// TIA Portal V15.1 export
// export: Created 2000-01-01T00:00:00.0000000Z, ExportSetting None
FUNCTION "FC_Rung" : Void   // FC42, LAD
{ S7_Optimized_Access := 'TRUE' }
   VAR_INPUT
      Local : Int;
   END_VAR
BEGIN

REGION Network 1
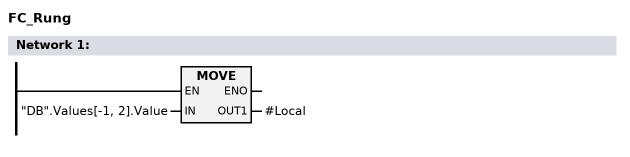
   RUNG wire#powerrail
      Move(in := "DB".Values[-1, 2].Value, out1 => #Local)
   END_RUNG
   // the same network as SCL:
   #Local := "DB".Values[-1, 2].Value;
END_REGION
END_FUNCTION
